(* IEC 61131-3 sources: com.logicals.npe.examples/HIS_Demo/.shadowcopy/src, 6 files *)

(* ---- FB_HISSafety.iecfbd ---- *)
(* Safety FBD template. Two equivalent NC contacts assumed.
   Requires the matching PLCopen Safety library and qualified HIS target setup.
   T#100ms is a DEMO PLACEHOLDER, not a validated discrepancy time.
   Safe communication loss must substitute FALSE at BOTH safe inputs.
   Never replace missing safe input data with standard BOOL simulation values.
   No auto reset or start reset. Reset does not start the process.
*)
FUNCTION_BLOCK FB_HISSafety
  USING safety.plcopen;
VAR_INPUT
    S_EStopA : SAFEBOOL;
    S_EStopB : SAFEBOOL;
    Reset : BOOL;
END_VAR
VAR_OUTPUT
    S_Permit : SAFEBOOL;
    SafetyDemand : BOOL;
    ResetRequest : BOOL;
    Error : BOOL;
    EquivalentDiag : WORD;
    EStopDiag : WORD;
END_VAR
VAR CONSTANT
    S_ResetDisabled : SAFEBOOL := FALSE;
END_VAR
VAR
    fbEquivalent : SF_Equivalent;
    fbEmergencyStop : SF_EmergencyStop;
END_VAR

  (*
    // Network 1: equivalent contacts, emergency stop, diagnostics
    fbEquivalent(Activate := TRUE, S_ChannelA := S_EStopA, S_ChannelB := S_EStopB, DiscrepancyTime := T#100ms);
    fbEmergencyStop(Activate := TRUE, S_EStopIn := fbEquivalent.S_EquivalentOut, S_StartReset := S_ResetDisabled, S_AutoReset := S_ResetDisabled, Reset := Reset, S_EStopOut => S_Permit, SafetyDemand => SafetyDemand, ResetRequest => ResetRequest, DiagCode => EStopDiag);
    EquivalentDiag := fbEquivalent.DiagCode;
    OR(IN1 := fbEquivalent.Error, IN2 := fbEmergencyStop.Error, OR => Error);
  *)

  @C(1) : @FB(fbEquivalent), @R(450.0, 90.0, 360.0, 194.0), @I(@N(Activate), @L(54.5)), @I(@N(S_ChannelA), @L(84.5)), @I(@N(S_ChannelB), @L(114.5)), @I(@N(DiscrepancyTime), @L(144.5)), @O(@N(Ready), @R(54.5)), @O(@N(S_EquivalentOut), @R(84.5)), @O(@N(SafetyDemand), @R(114.5)), @O(@N(Error), @R(144.5)), @O(@N(DiagCode), @R(174.5));
  @C(2) : @FB(fbEmergencyStop), @R(1260.0, 90.0, 360.0, 224.0), @I(@N(Activate), @L(54.5)), @I(@N(S_EStopIn), @L(84.5)), @I(@N(S_StartReset), @L(114.5)), @I(@N(S_AutoReset), @L(144.5)), @I(@N(Reset), @L(174.5)), @O(@N(Ready), @R(54.5)), @O(@N(S_EStopOut), @R(84.5)), @O(@N(SafetyDemand), @R(114.5)), @O(@N(ResetRequest), @R(144.5)), @O(@N(Error), @R(174.5)), @O(@N(DiagCode), @R(204.5));
  @VF(3) : @E(S_EStopA), @R(45.0, 165.0, 300.0, 19.0);
  @VF(4) : @E(S_EStopB), @R(45.0, 195.0, 300.0, 19.0);
  @VF(5) : @E(Reset), @R(870.0, 255.0, 300.0, 19.0);
  @VF(6) : @E(S_Permit), @R(1710.0, 165.0, 300.0, 19.0);
  @VF(7) : @E(SafetyDemand), @R(1710.0, 195.0, 300.0, 19.0);
  @VF(8) : @E(ResetRequest), @R(1710.0, 225.0, 300.0, 19.0);
  @VF(9) : @E(EStopDiag), @R(1710.0, 285.0, 300.0, 19.0);
  @VF(10) : @E(EquivalentDiag), @R(870.0, 375.0, 300.0, 19.0);
  @C(11) : @F(OR), @R(1260.0, 510.0, 180.0, 104.0), BOOL, @I(@N(IN1), @L(54.5)), @I(@N(IN2), @L(84.5)), @O(@N(OR), @R(54.5));
  @VF(12) : @E(Error), @R(1530.0, 555.0, 300.0, 19.0);

  @VF(25) : @E(TRUE), @R(45.0, 135.0, 300.0, 19.0);
  @VF(26) : @E(T#100ms), @R(45.0, 225.0, 300.0, 19.0);
  @VF(27) : @E(TRUE), @R(870.0, 135.0, 300.0, 19.0);
  @VF(28) : @E(S_ResetDisabled), @R(870.0, 195.0, 300.0, 19.0);
  @VF(29) : @E(S_ResetDisabled), @R(870.0, 225.0, 300.0, 19.0);

  @G(13) : @L(@VF(3).o, @C(1).S_ChannelA);
  @G(14) : @L(@VF(4).o, @C(1).S_ChannelB);
  @G(15) : @L(@C(1).S_EquivalentOut, @C(2).S_EStopIn);
  @G(16) : @L(@VF(5).o, @C(2).Reset);
  @G(17) : @L(@C(2).S_EStopOut, @VF(6).i);
  @G(18) : @L(@C(2).SafetyDemand, @VF(7).i);
  @G(19) : @L(@C(2).ResetRequest, @VF(8).i);
  @G(20) : @L(@C(2).DiagCode, @VF(9).i);
  @G(21) : @L(@C(1).DiagCode, @VF(10).i);
  @G(22) : @L(@C(1).Error, @C(11).IN1);
  @G(23) : @L(@C(2).Error, @C(11).IN2);
  @G(24) : @L(@C(11).OR, @VF(12).i);
  @G(30) : @L(@VF(25).o, @C(1).Activate);
  @G(31) : @L(@VF(26).o, @C(1).DiscrepancyTime);
  @G(32) : @L(@VF(27).o, @C(2).Activate);
  @G(33) : @L(@VF(28).o, @C(2).S_StartReset);
  @G(34) : @L(@VF(29).o, @C(2).S_AutoReset);
END_FUNCTION_BLOCK

(* ---- FB_PackagingDataSimulation.iecst ---- *)
(* Simulation-only synthetic process data and harmless demo-load outputs.
 * Called after FB_PackagingLine, only in SimMode. Not a safety function.
 *)
FUNCTION_BLOCK FB_PackagingDataSimulation
    VAR_INPUT
        Reset : BOOL;
        S_Permit : SAFEBOOL;
        S_EStopReleased : SAFEBOOL;
        LineState : UINT;
        LineFault : BOOL;
        CycleDone : BOOL;
        FastCycle : BOOL;
        Heartbeat : BOOL;
    END_VAR
    VAR_OUTPUT
        S_DataPlausible : SAFEBOOL;
    END_VAR
    VAR
        tSecond : TON;
        PrevJam : BOOL;
        PrevGuardClosed : SAFEBOOL := TRUE;
        PrevEStopReleased : SAFEBOOL := FALSE;
        PreviousLineState : UINT;
    END_VAR
    VAR_EXTERNAL
        S_InfeedGuardClosed : SAFEBOOL;
        S_SealingGuardClosed : SAFEBOOL;
        S_OutfeedGuardClosed : SAFEBOOL;
        S_ServiceDoorClosed : SAFEBOOL;
        S_AirSupplyReady : SAFEBOOL;
        S_InfeedZoneStatus : SAFEBYTE;
        S_SealingZoneStatus : SAFEBYTE;
        S_OutfeedZoneStatus : SAFEBYTE;
        S_GuardLockStatus : SAFEBYTE;
        S_SafeDriveStatus : SAFEBYTE;
        S_InfeedDiagnosticCode : SAFEWORD;
        S_SealingDiagnosticCode : SAFEWORD;
        S_OutfeedDiagnosticCode : SAFEWORD;
        S_SafetyBusDiagnosticCode : SAFEWORD;
        S_DriveDiagnosticCode : SAFEWORD;
        S_ZonePermissionMask : SAFEDWORD;
        S_GuardMonitoringMask : SAFEDWORD;
        S_DriveEnableMask : SAFEDWORD;
        S_ActiveSafetyDemandMask : SAFEDWORD;
        S_ConfirmedSafetyDemandMask : SAFEDWORD;
        S_InfeedMotionDirection : SAFESINT;
        S_SealingMotionDirection : SAFESINT;
        S_OutfeedMotionDirection : SAFESINT;
        S_FilmFeedMotionDirection : SAFESINT;
        S_RejectGateMotionDirection : SAFESINT;
        S_SealingTemperatureLimit_dC : SAFEINT;
        S_SealingTemperatureActual_dC : SAFEINT;
        S_AmbientTemperatureActual_dC : SAFEINT;
        S_MinSealingTemperature_dC : SAFEINT;
        S_MaxSealingTemperature_dC : SAFEINT;
        S_InfeedStopPosition_mm : SAFEDINT;
        S_SealingStopPosition_mm : SAFEDINT;
        S_OutfeedStopPosition_mm : SAFEDINT;
        S_CartonTrackingPosition_mm : SAFEDINT;
        S_MaxStoppingDistance_mm : SAFEDINT;
        S_InfeedSensorCount : SAFEUSINT;
        S_SealingSensorCount : SAFEUSINT;
        S_OutfeedSensorCount : SAFEUSINT;
        S_GuardChannelCount : SAFEUSINT;
        S_DriveFeedbackChannelCount : SAFEUSINT;
        S_InfeedSpeedLimit_mm_s : SAFEUINT;
        S_OutfeedSpeedLimit_mm_s : SAFEUINT;
        S_MinAirPressure_mbar : SAFEUINT;
        S_MaxAirPressure_mbar : SAFEUINT;
        S_MotorCurrentLimit_mA : SAFEUINT;
        S_CompletedCartonCount : SAFEUDINT;
        S_RejectedCartonCount : SAFEUDINT;
        S_GuardOpeningCount : SAFEUDINT;
        S_EStopDemandCount : SAFEUDINT;
        S_OperatingTime_s : SAFEUDINT;
        O01 : BOOL;
        O02 : BOOL;
        O03 : BOOL;
        O04 : BOOL;
        O14 : BOOL;
        O15 : BOOL;
        O16 : BOOL;
        O17 : BOOL;
        O18 : BOOL;
        SO01 : SAFEBOOL;
        SO02 : SAFEBOOL;
        SO12 : SAFEBOOL;
        SO13 : SAFEBOOL;
        SO14 : SAFEBOOL;
    END_VAR

    IF Reset THEN
        S_CompletedCartonCount := 0;
        S_RejectedCartonCount := 0;
        S_GuardOpeningCount := 0;
        S_EStopDemandCount := 0;
        S_OperatingTime_s := 0;
        S_SealingTemperatureActual_dC := 1650;
        S_CartonTrackingPosition_mm := 0;
        PrevJam := LineFault;
        PrevGuardClosed := TRUE;
        PrevEStopReleased := S_EStopReleased;
        PreviousLineState := 0;
    END_IF;
    (* Telemetry tick: task-quantised nominal second, not a precision clock. *)
    tSecond(IN := NOT tSecond.Q AND NOT Reset, PT := T#1s);

    S_InfeedGuardClosed := TRUE;
    S_SealingGuardClosed := TRUE;
    S_OutfeedGuardClosed := TRUE;
    S_ServiceDoorClosed := TRUE;
    IF LineFault THEN S_ServiceDoorClosed := FALSE; END_IF;
    S_AirSupplyReady := S_EStopReleased;
    S_SealingTemperatureLimit_dC := 1800;
    S_MinSealingTemperature_dC := 1600;
    S_MaxSealingTemperature_dC := 2000;
    S_AmbientTemperatureActual_dC := 230;
    S_InfeedStopPosition_mm := 1000;
    S_SealingStopPosition_mm := 2000;
    S_OutfeedStopPosition_mm := 3000;
    S_MaxStoppingDistance_mm := 200;
    S_InfeedSpeedLimit_mm_s := 250;
    S_OutfeedSpeedLimit_mm_s := 250;
    IF FastCycle THEN
        S_InfeedSpeedLimit_mm_s := 500;
        S_OutfeedSpeedLimit_mm_s := 500;
    END_IF;
    S_MinAirPressure_mbar := 5500;
    S_MaxAirPressure_mbar := 7500;
    S_MotorCurrentLimit_mA := 4500;
    S_InfeedSensorCount := 2;
    S_SealingSensorCount := 2;
    S_OutfeedSensorCount := 2;
    S_GuardChannelCount := 4;
    S_DriveFeedbackChannelCount := 3;

    (* Zone status 0 blocked, 1 idle, 2 moving, 3 jam. *)
    S_InfeedZoneStatus := 0;
    S_SealingZoneStatus := 0;
    S_OutfeedZoneStatus := 0;
    IF S_Permit AND NOT LineFault THEN
        S_InfeedZoneStatus := 1;
        S_SealingZoneStatus := 1;
        S_OutfeedZoneStatus := 1;
        IF LineState = 20 THEN S_InfeedZoneStatus := 2; END_IF;
        IF LineState = 30 THEN S_SealingZoneStatus := 2; END_IF;
        IF LineState = 40 THEN S_OutfeedZoneStatus := 2; END_IF;
    END_IF;
    IF LineFault THEN S_SealingZoneStatus := 3; END_IF;
    S_GuardLockStatus := 1;
    IF NOT S_ServiceDoorClosed THEN S_GuardLockStatus := 0; END_IF;
    S_SafeDriveStatus := 0;
    IF S_Permit AND S_ServiceDoorClosed THEN S_SafeDriveStatus := 1; END_IF;
    S_InfeedDiagnosticCode := 0;
    S_SealingDiagnosticCode := 0;
    S_OutfeedDiagnosticCode := 0;
    S_SafetyBusDiagnosticCode := 0;
    S_DriveDiagnosticCode := 0;
    IF LineFault THEN S_SealingDiagnosticCode := 16#1001; END_IF;
    IF NOT S_EStopReleased THEN S_SafetyBusDiagnosticCode := 16#2001; END_IF;
    IF NOT S_Permit THEN S_DriveDiagnosticCode := 16#3001; END_IF;

    (* Zones bits 0..2, guards bits 0..3; demand bit 0 E-stop,
       bit 1 virtual service access during jam recovery. *)
    S_ZonePermissionMask := 0;
    IF S_Permit AND S_ServiceDoorClosed AND S_AirSupplyReady THEN S_ZonePermissionMask := 7; END_IF;
    S_GuardMonitoringMask := 15;
    IF NOT S_ServiceDoorClosed THEN S_GuardMonitoringMask := 7; END_IF;
    (* SAFEDWORD is a bitstring, not an arithmetic integer.
       Explicit patterns: bit 0 = E-stop, bit 1 = virtual service door. *)
    S_ActiveSafetyDemandMask := 16#00000000;
    IF NOT S_EStopReleased THEN
        S_ActiveSafetyDemandMask := 16#00000001;
        IF NOT S_ServiceDoorClosed THEN S_ActiveSafetyDemandMask := 16#00000003; END_IF;
    ELSIF NOT S_ServiceDoorClosed THEN
        S_ActiveSafetyDemandMask := 16#00000002;
    END_IF;
    S_ConfirmedSafetyDemandMask := S_ActiveSafetyDemandMask;
    S_DriveEnableMask := 0;
    S_InfeedMotionDirection := 0;
    S_SealingMotionDirection := 0;
    S_OutfeedMotionDirection := 0;
    S_FilmFeedMotionDirection := 0;
    S_RejectGateMotionDirection := 0;
    IF S_ZonePermissionMask = 7 THEN
        IF LineState = 20 THEN S_DriveEnableMask := 1; S_InfeedMotionDirection := 1; END_IF;
        IF LineState = 30 THEN S_DriveEnableMask := 2; S_SealingMotionDirection := 1; S_FilmFeedMotionDirection := 1; END_IF;
        IF LineState = 40 THEN S_DriveEnableMask := 4; S_OutfeedMotionDirection := 1; END_IF;
    END_IF;
    (* Signed virtual sample; no physical motor is commanded in reverse. *)
    IF LineFault THEN S_RejectGateMotionDirection := -1; END_IF;

    IF LineState <> PreviousLineState THEN
        IF LineState = 20 THEN S_CartonTrackingPosition_mm := 0; END_IF;
        IF (LineState = 30) OR (LineState = 40) THEN S_CartonTrackingPosition_mm := S_SealingStopPosition_mm; END_IF;
        IF LineState = 50 THEN S_CartonTrackingPosition_mm := S_OutfeedStopPosition_mm; END_IF;
    END_IF;
    IF (LineState = 0) OR (LineState = 10) THEN S_CartonTrackingPosition_mm := 0; END_IF;
    IF tSecond.Q THEN
        IF S_OperatingTime_s < 1000000000 THEN S_OperatingTime_s := S_OperatingTime_s + 1; END_IF;
        IF S_SealingTemperatureActual_dC < S_SealingTemperatureLimit_dC THEN
            S_SealingTemperatureActual_dC := S_SealingTemperatureActual_dC + 10;
            IF S_SealingTemperatureActual_dC > S_SealingTemperatureLimit_dC THEN S_SealingTemperatureActual_dC := S_SealingTemperatureLimit_dC; END_IF;
        END_IF;
        IF (S_InfeedMotionDirection = 1) AND (S_CartonTrackingPosition_mm < S_InfeedStopPosition_mm) THEN
            S_CartonTrackingPosition_mm := S_CartonTrackingPosition_mm + 250;
            IF S_CartonTrackingPosition_mm > S_InfeedStopPosition_mm THEN S_CartonTrackingPosition_mm := S_InfeedStopPosition_mm; END_IF;
        END_IF;
        IF (S_OutfeedMotionDirection = 1) AND (S_CartonTrackingPosition_mm < S_OutfeedStopPosition_mm) THEN
            S_CartonTrackingPosition_mm := S_CartonTrackingPosition_mm + 250;
            IF S_CartonTrackingPosition_mm > S_OutfeedStopPosition_mm THEN S_CartonTrackingPosition_mm := S_OutfeedStopPosition_mm; END_IF;
        END_IF;
    END_IF;
    (* Separate simulation-session counters, saturated rather than wrapped. *)
    IF NOT Reset THEN
        IF CycleDone AND (S_CompletedCartonCount < 1000000000) THEN S_CompletedCartonCount := S_CompletedCartonCount + 1; END_IF;
        IF LineFault AND NOT PrevJam AND (S_RejectedCartonCount < 1000000000) THEN S_RejectedCartonCount := S_RejectedCartonCount + 1; END_IF;
        IF NOT S_ServiceDoorClosed AND PrevGuardClosed AND (S_GuardOpeningCount < 1000000000) THEN S_GuardOpeningCount := S_GuardOpeningCount + 1; END_IF;
        IF NOT S_EStopReleased AND PrevEStopReleased AND (S_EStopDemandCount < 1000000000) THEN S_EStopDemandCount := S_EStopDemandCount + 1; END_IF;
    END_IF;
    PrevJam := LineFault;
    PrevGuardClosed := S_ServiceDoorClosed;
    PrevEStopReleased := S_EStopReleased;
    PreviousLineState := LineState;

    (* All 50 globals are read in the validity/data chain below. *)
    S_DataPlausible :=
        S_InfeedGuardClosed AND S_SealingGuardClosed AND S_OutfeedGuardClosed
        AND (S_ServiceDoorClosed OR (S_GuardLockStatus = 0))
        AND (S_AirSupplyReady OR (S_ActiveSafetyDemandMask <> 0))
        AND (S_InfeedZoneStatus <= 3) AND (S_SealingZoneStatus <= 3) AND (S_OutfeedZoneStatus <= 3)
        AND (S_GuardLockStatus <= 1) AND (S_SafeDriveStatus <= 1)
        AND (S_InfeedDiagnosticCode = 0) AND ((S_SealingDiagnosticCode = 0) OR (S_SealingDiagnosticCode = 16#1001))
        AND (S_OutfeedDiagnosticCode = 0) AND ((S_SafetyBusDiagnosticCode = 0) OR (S_SafetyBusDiagnosticCode = 16#2001))
        AND ((S_DriveDiagnosticCode = 0) OR (S_DriveDiagnosticCode = 16#3001))
        AND (S_ZonePermissionMask <= 7) AND (S_GuardMonitoringMask <= 15) AND (S_DriveEnableMask <= 7)
        AND (S_ActiveSafetyDemandMask <= 3) AND (S_ConfirmedSafetyDemandMask = S_ActiveSafetyDemandMask)
        AND (S_InfeedMotionDirection >= 0) AND (S_InfeedMotionDirection <= 1)
        AND (S_SealingMotionDirection >= 0) AND (S_SealingMotionDirection <= 1)
        AND (S_OutfeedMotionDirection >= 0) AND (S_OutfeedMotionDirection <= 1)
        AND (S_FilmFeedMotionDirection >= 0) AND (S_FilmFeedMotionDirection <= 1)
        AND (S_RejectGateMotionDirection >= -1) AND (S_RejectGateMotionDirection <= 0)
        AND (S_SealingTemperatureLimit_dC >= S_MinSealingTemperature_dC)
        AND (S_SealingTemperatureLimit_dC <= S_MaxSealingTemperature_dC)
        AND (S_SealingTemperatureActual_dC >= S_MinSealingTemperature_dC)
        AND (S_SealingTemperatureActual_dC <= S_MaxSealingTemperature_dC)
        AND (S_AmbientTemperatureActual_dC >= 0) AND (S_AmbientTemperatureActual_dC <= 500)
        AND (S_InfeedStopPosition_mm > S_MaxStoppingDistance_mm)
        AND (S_SealingStopPosition_mm > S_InfeedStopPosition_mm)
        AND (S_OutfeedStopPosition_mm > S_SealingStopPosition_mm)
        AND (S_CartonTrackingPosition_mm >= 0) AND (S_CartonTrackingPosition_mm <= S_OutfeedStopPosition_mm)
        AND (S_InfeedSensorCount = 2) AND (S_SealingSensorCount = 2) AND (S_OutfeedSensorCount = 2)
        AND (S_GuardChannelCount = 4) AND (S_DriveFeedbackChannelCount = 3)
        AND (S_InfeedSpeedLimit_mm_s > 0) AND (S_InfeedSpeedLimit_mm_s <= 500)
        AND (S_OutfeedSpeedLimit_mm_s > 0) AND (S_OutfeedSpeedLimit_mm_s <= 500)
        AND (S_MinAirPressure_mbar < S_MaxAirPressure_mbar) AND (S_MotorCurrentLimit_mA > 0)
        AND (S_CompletedCartonCount <= 1000000000) AND (S_RejectedCartonCount <= 1000000000)
        AND (S_GuardOpeningCount = S_RejectedCartonCount)
        AND (S_EStopDemandCount <= 1000000000) AND (S_OperatingTime_s <= 1000000000);

    O01 := S_Permit AND S_DataPlausible AND (S_InfeedMotionDirection = 1);
    O02 := S_Permit AND S_DataPlausible AND (S_SealingMotionDirection = 1);
    O03 := S_Permit AND S_DataPlausible AND (S_OutfeedMotionDirection = 1);
    O04 := S_Permit AND S_DataPlausible AND (S_FilmFeedMotionDirection = 1);
    O14 := S_Permit AND S_DataPlausible AND (S_ZonePermissionMask = 7);
    O15 := S_Permit AND S_DataPlausible AND Heartbeat;
    O16 := S_Permit AND S_DataPlausible AND (S_SealingDiagnosticCode <> 0);
    O17 := S_Permit AND S_DataPlausible AND (S_SealingTemperatureActual_dC >= S_SealingTemperatureLimit_dC);
    O18 := S_Permit AND S_DataPlausible AND (S_GuardMonitoringMask = 15);
    (* Safe-typed expressions; demo indications, not validated safety outputs. *)
    SO01 := S_Permit AND S_DataPlausible AND S_AirSupplyReady;
    SO02 := S_Permit AND S_DataPlausible AND S_ServiceDoorClosed;
    SO12 := S_Permit AND S_DataPlausible AND S_InfeedGuardClosed AND (S_InfeedMotionDirection = 1);
    SO13 := S_Permit AND S_DataPlausible AND S_SealingGuardClosed AND (S_SealingMotionDirection = 1);
    SO14 := S_Permit AND S_DataPlausible AND S_OutfeedGuardClosed AND (S_OutfeedMotionDirection = 1);
END_FUNCTION_BLOCK

(* ---- FB_PackagingIndicators.iecfbd ---- *)
(* Non-safety FBD. Suggested four standard LED functions.
   All physical output assignments remain open.
*)
FUNCTION_BLOCK FB_PackagingIndicators
VAR_INPUT
    Permit : BOOL;
    Ready : BOOL;
    Infeed : BOOL;
    Sealing : BOOL;
    Outfeed : BOOL;
    Complete : BOOL;
    Blocked : BOOL;
    ProcessFault : BOOL;
    SafetyError : BOOL;
    ResetRequest : BOOL;
    Heartbeat : BOOL;
END_VAR
VAR_OUTPUT
    LedReady : BOOL;
    LedConveyor : BOOL;
    LedSealing : BOOL;
    LedAttention : BOOL;
END_VAR

  (*
    Explicit Boolean gates; value fields contain single variables only.
    OR(IN1 := Ready, IN2 := Complete);
    AND(IN1 := Permit, IN2 := @C(1).OR);
    OR(IN1 := Infeed, IN2 := Outfeed);
    AND(IN1 := Permit, IN2 := @C(7).OR, IN3 := Heartbeat);
    AND(IN1 := Permit, IN2 := Sealing, IN3 := Heartbeat);
    NOT(IN := ResetRequest);
    AND(IN1 := Blocked, IN2 := @C(19).NOT);
    AND(IN1 := ResetRequest, IN2 := Heartbeat);
    OR(IN1 := @C(21).AND, IN2 := ProcessFault, IN3 := SafetyError, IN4 := @C(23).AND);
  *)

  @C(1) : @F(OR), @R(390.0, 90.0, 180.0, 104.0), BOOL, @I(@N(IN1), @L(54.5)), @I(@N(IN2), @L(84.5)), @O(@N(OR), @R(54.5));
  @VF(2) : @E(Ready), @R(45.0, 135.0, 180.0, 19.0);
  @VF(3) : @E(Complete), @R(45.0, 165.0, 180.0, 19.0);
  @C(4) : @F(AND), @R(900.0, 60.0, 180.0, 104.0), BOOL, @I(@N(IN1), @L(54.5)), @I(@N(IN2), @L(84.5)), @O(@N(AND), @R(54.5));
  @VF(5) : @E(Permit), @R(645.0, 105.0, 180.0, 19.0);
  @VF(6) : @E(LedReady), @R(1230.0, 105.0, 180.0, 19.0);
  @C(7) : @F(OR), @R(390.0, 390.0, 180.0, 104.0), BOOL, @I(@N(IN1), @L(54.5)), @I(@N(IN2), @L(84.5)), @O(@N(OR), @R(54.5));
  @VF(8) : @E(Infeed), @R(45.0, 435.0, 180.0, 19.0);
  @VF(9) : @E(Outfeed), @R(45.0, 465.0, 180.0, 19.0);
  @C(10) : @F(AND), @R(900.0, 360.0, 180.0, 134.0), BOOL, @I(@N(IN1), @L(54.5)), @I(@N(IN2), @L(84.5)), @I(@N(IN3), @L(114.5)), @O(@N(AND), @R(54.5));
  @VF(11) : @E(Permit), @R(645.0, 405.0, 180.0, 19.0);
  @VF(12) : @E(Heartbeat), @R(645.0, 465.0, 180.0, 19.0);
  @VF(13) : @E(LedConveyor), @R(1230.0, 405.0, 180.0, 19.0);
  @C(14) : @F(AND), @R(900.0, 660.0, 180.0, 134.0), BOOL, @I(@N(IN1), @L(54.5)), @I(@N(IN2), @L(84.5)), @I(@N(IN3), @L(114.5)), @O(@N(AND), @R(54.5));
  @VF(15) : @E(Permit), @R(645.0, 705.0, 180.0, 19.0);
  @VF(16) : @E(Sealing), @R(645.0, 735.0, 180.0, 19.0);
  @VF(17) : @E(Heartbeat), @R(645.0, 765.0, 180.0, 19.0);
  @VF(18) : @E(LedSealing), @R(1230.0, 705.0, 180.0, 19.0);
  @C(19) : @F(NOT), @R(375.0, 1080.0, 180.0, 74.0), BOOL, @I(@N(IN), @L(54.5)), @O(@N(NOT), @R(54.5));
  @VF(20) : @E(ResetRequest), @R(45.0, 1125.0, 180.0, 19.0);
  @C(21) : @F(AND), @R(660.0, 1050.0, 180.0, 104.0), BOOL, @I(@N(IN1), @L(54.5)), @I(@N(IN2), @L(84.5)), @O(@N(AND), @R(54.5));
  @VF(22) : @E(Blocked), @R(375.0, 1035.0, 180.0, 19.0);
  @C(23) : @F(AND), @R(660.0, 1230.0, 180.0, 104.0), BOOL, @I(@N(IN1), @L(54.5)), @I(@N(IN2), @L(84.5)), @O(@N(AND), @R(54.5));
  @VF(24) : @E(ResetRequest), @R(375.0, 1275.0, 180.0, 19.0);
  @VF(25) : @E(Heartbeat), @R(375.0, 1305.0, 180.0, 19.0);
  @C(26) : @F(OR), @R(1200.0, 1050.0, 180.0, 164.0), BOOL, @I(@N(IN1), @L(54.5)), @I(@N(IN2), @L(84.5)), @I(@N(IN3), @L(114.5)), @I(@N(IN4), @L(144.5)), @O(@N(OR), @R(54.5));
  @VF(27) : @E(ProcessFault), @R(930.0, 1125.0, 180.0, 19.0);
  @VF(28) : @E(SafetyError), @R(930.0, 1155.0, 180.0, 19.0);
  @VF(29) : @E(LedAttention), @R(1500.0, 1095.0, 180.0, 19.0);

  @G(30) : @L(@VF(2).o, @C(1).IN1);
  @G(31) : @L(@VF(3).o, @C(1).IN2);
  @G(32) : @L(@VF(5).o, @C(4).IN1);
  @G(33) : @L(@C(1).OR, @C(4).IN2);
  @G(34) : @L(@C(4).AND, @VF(6).i);
  @G(35) : @L(@VF(8).o, @C(7).IN1);
  @G(36) : @L(@VF(9).o, @C(7).IN2);
  @G(37) : @L(@VF(11).o, @C(10).IN1);
  @G(38) : @L(@C(7).OR, @C(10).IN2);
  @G(39) : @L(@VF(12).o, @C(10).IN3);
  @G(40) : @L(@C(10).AND, @VF(13).i);
  @G(41) : @L(@VF(15).o, @C(14).IN1);
  @G(42) : @L(@VF(16).o, @C(14).IN2);
  @G(43) : @L(@VF(17).o, @C(14).IN3);
  @G(44) : @L(@C(14).AND, @VF(18).i);
  @G(45) : @L(@VF(20).o, @C(19).IN);
  @G(46) : @L(@VF(22).o, @C(21).IN1);
  @G(47) : @L(@C(19).NOT, @C(21).IN2);
  @G(48) : @L(@VF(24).o, @C(23).IN1);
  @G(49) : @L(@VF(25).o, @C(23).IN2);
  @G(50) : @L(@C(21).AND, @C(26).IN1);
  @G(51) : @L(@VF(27).o, @C(26).IN2);
  @G(52) : @L(@VF(28).o, @C(26).IN3);
  @G(53) : @L(@C(23).AND, @C(26).IN4);
  @G(54) : @L(@C(26).OR, @VF(29).i);
END_FUNCTION_BLOCK

(* ---- FB_PackagingLine.iecst ---- *)
(* HIS Packaging Line / SPS 2026
 *    Non-safety simulation. Never use these outputs as a safety function.
 *    Call once per cyclic task. No physical I/O addresses are assigned.
 *)
FUNCTION_BLOCK FB_PackagingLine
	VAR_INPUT
		Enable : BOOL;
		Permit : BOOL; (* Read-only status copy from the safety POU. *)
		Start : BOOL;
		Stop : BOOL;
		FastCycle : BOOL;
		Jam : BOOL; (* Simulated carton jam, NOT a safety fault. *)
		AckJam : BOOL;
	END_VAR
	VAR_OUTPUT
		State : UINT;
		(* 0 blocked, 10 ready, 20 infeed, 30 sealing,
		 40 outfeed, 50 complete, 90 carton jam *)
		Ready : BOOL;
		Infeed : BOOL;
		Sealing : BOOL;
		Outfeed : BOOL;
		Complete : BOOL;
		Blocked : BOOL;
		Fault : BOOL;
		Running : BOOL;
		Heartbeat : BOOL;
		CycleDone : BOOL; (* One scan pulse after carton leaves station. *)
		CartonsPacked : UDINT;
		FastCycleActive : BOOL;
	END_VAR
	VAR
		PrevStart : BOOL;
		PrevAck : BOOL;
		FirstScan : BOOL := TRUE;
		StartEdge : BOOL;
		AckEdge : BOOL;
		StartArmed : BOOL;
		FaultLatched : BOOL;
		InfeedTime : TIME := T#3s;
		SealTime : TIME := T#2s;
		OutfeedTime : TIME := T#2s;
		tInfeed : TON;
		tSeal : TON;
		tOutfeed : TON;
		tSuccess : TON;
		tBlink : TON;
	END_VAR

	(* Suppress edges on startup; held Start never causes a restart. *)
	StartEdge := Start AND NOT PrevStart AND NOT FirstScan;
	AckEdge := AckJam AND NOT PrevAck AND NOT FirstScan;
	PrevStart := Start;
	PrevAck := AckJam;
	FirstScan := FALSE;
	CycleDone := FALSE;

	(* Timers are executed on every scan, also when disabled. *)
	tBlink(IN := NOT tBlink.Q, PT := T#250ms);
	IF tBlink.Q THEN
		Heartbeat := NOT Heartbeat;
	END_IF;
	tInfeed(IN := (State = 20) AND Enable AND Permit AND NOT Stop
            AND NOT Jam, PT := InfeedTime);
	tSeal(IN := (State = 30) AND Enable AND Permit AND NOT Stop
             AND NOT Jam, PT := SealTime);
	tOutfeed(IN := (State = 40) AND Enable AND Permit AND NOT Stop
              AND NOT Jam, PT := OutfeedTime);
	tSuccess(IN := (State = 50) AND Enable AND Permit AND NOT Stop
               AND NOT Jam, PT := T#1s);

	(* Keep process faults latched even across a safety interruption. *)
	IF Jam AND Enable AND Permit
   AND ((State = 20) OR (State = 30) OR (State = 40)) THEN
		FaultLatched := TRUE;
	END_IF;
	IF AckEdge AND NOT Jam AND Enable AND Permit THEN
		FaultLatched := FALSE;
	END_IF;

	(* Priority: no permit / disabled > process fault > stop > sequence. *)
	IF NOT Enable OR NOT Permit THEN
		State := 0;

		FastCycleActive := FALSE;
		StartArmed := FALSE;
	ELSIF FaultLatched THEN
		State := 90;

		FastCycleActive := FALSE;
		StartArmed := FALSE;
	ELSIF Stop THEN
		State := 10;

		FastCycleActive := FALSE;
		StartArmed := FALSE;
	ELSE
		CASE State OF
			0, 90:
			State := 10;

			FastCycleActive := FALSE;
			StartArmed := FALSE;
			10:
            IF NOT Start THEN
				StartArmed := TRUE;
			END_IF;
			IF StartEdge AND StartArmed AND NOT Jam
               AND NOT AckJam THEN
				FastCycleActive := FastCycle; (* Latch throughput mode for this carton. *)
				IF FastCycleActive THEN
					InfeedTime := T#1500ms;
					SealTime := T#1s;
					OutfeedTime := T#1s;
				ELSE
					InfeedTime := T#3s;
					SealTime := T#2s;
					OutfeedTime := T#2s;
				END_IF;
				StartArmed := FALSE;

				State := 20;
			END_IF;
			20:
            IF tInfeed.Q THEN
				State := 30;
			END_IF;
			30:
            IF tSeal.Q THEN

				State := 40;
			END_IF;
			40:
            IF tOutfeed.Q THEN
				IF CartonsPacked < UDINT#4294967295 THEN
					CartonsPacked := CartonsPacked + 1;
				END_IF;
				CycleDone := TRUE;
				State := 50;
			END_IF;
			50:
            IF tSuccess.Q THEN
				State := 10;
				FastCycleActive := FALSE;
				StartArmed := FALSE;
			END_IF;
		ELSE
			FaultLatched := TRUE;
			State := 90;

			FastCycleActive := FALSE;
			StartArmed := FALSE;
		END_CASE;
	END_IF;

	Blocked := NOT Enable OR NOT Permit;
	Fault := FaultLatched;
	Ready := (State = 10) AND Enable AND Permit AND NOT FaultLatched
         AND NOT Stop AND NOT Jam AND NOT AckJam;
	Infeed := State = 20;
	Sealing := State = 30;
	Outfeed := State = 40;
	Complete := State = 50;
	Running := Infeed OR Sealing OR Outfeed;
END_FUNCTION_BLOCK

(* ---- FB_PackagingSimulation.iecst ---- *)
(* Automatic exhibition simulation; not a physical safety input source.
 * Called ONLY while PRG_HISDemo.SimMode is TRUE.
 * Drives simulated commands through the unchanged safety/process blocks.
 * Reset on every mode entry; feedback comes from the previous program scan.
 *)
FUNCTION_BLOCK FB_PackagingSimulation
    VAR_INPUT
        Reset : BOOL;
        Permit : BOOL;
        LineReady : BOOL;
        LineState : UINT;
        LineFault : BOOL;
        InjectFaults : BOOL;
        FastCycle : BOOL;
    END_VAR
    VAR_OUTPUT
        EStopReleased : SAFEBOOL;
        Enable : BOOL;
        Start : BOOL;
        Stop : BOOL;
        SafetyReset : BOOL;
        Jam : BOOL;
        AckJam : BOOL;
        FastCycleCommand : BOOL;
        (* 0 boot; 10 release; 20 reset gap; 30 reset pulse; 40 ready;
           50 start pulse; 60 packaging; 70 jam; 80 clear jam;
           90 acknowledge; 100 emergency stop. *)
        State : UINT;
        AttemptInRound : UINT;
        (* 0 none; 1 normal carton; 2 jam demonstration; 3 E-stop demonstration. *)
        Scenario : UINT;
    END_VAR
    VAR
        tBoot : TON;
        tRelease : TON;
        tResetGap : TON;
        tResetPulse : TON;
        tReady : TON;
        tStart : TON;
        tJam : TON;
        tJamClear : TON;
        tAck : TON;
        tEStop : TON;
    END_VAR

    IF Reset THEN
        State := 0;
        AttemptInRound := 0;
        Scenario := 0;
    END_IF;

    (* Separate timers ensure every phase receives a fresh interval.
       Reset also clears timers left active when the block was not called. *)
    tBoot(IN := (State = 0) AND NOT Reset, PT := T#1s);
    tRelease(IN := (State = 10) AND NOT Reset, PT := T#1s);
    tResetGap(IN := (State = 20) AND NOT Reset, PT := T#500ms);
    tResetPulse(IN := (State = 30) AND NOT Reset, PT := T#500ms);
    tReady(IN := (State = 40) AND LineReady AND Permit AND NOT Reset, PT := T#500ms);
    tStart(IN := (State = 50) AND NOT Reset, PT := T#500ms);
    tJam(IN := (State = 70) AND NOT Reset, PT := T#3s);
    tJamClear(IN := (State = 80) AND NOT Reset, PT := T#500ms);
    tAck(IN := (State = 90) AND NOT Reset, PT := T#500ms);
    tEStop(IN := (State = 100) AND NOT Reset, PT := T#3s);

    IF NOT Reset THEN
        CASE State OF
            0:
                IF tBoot.Q THEN State := 10; END_IF;
            10:
                IF tRelease.Q THEN State := 20; END_IF;
            20:
                IF Permit THEN
                    IF LineFault THEN State := 80; ELSE State := 40; END_IF;
                ELSIF tResetGap.Q THEN
                    State := 30;
                END_IF;
            30:
                IF tResetPulse.Q THEN
                    IF Permit THEN
                        IF LineFault THEN State := 80; ELSE State := 40; END_IF;
                    ELSE
                        State := 20;
                    END_IF;
                END_IF;
            40:
                IF NOT Permit THEN
                    State := 10;
                ELSIF LineFault THEN
                    State := 80;
                ELSIF tReady.Q THEN
                    IF AttemptInRound >= 6 THEN AttemptInRound := 0; END_IF;
                    AttemptInRound := AttemptInRound + 1;
                    Scenario := 1;
                    IF InjectFaults AND (AttemptInRound = 3) THEN Scenario := 2; END_IF;
                    IF InjectFaults AND (AttemptInRound = 6) THEN Scenario := 3; END_IF;
                    State := 50;
                END_IF;
            50:
                IF NOT Permit THEN
                    State := 10;
                ELSIF tStart.Q THEN
                    State := 60;
                END_IF;
            60:
                IF NOT Permit THEN
                    State := 10;
                ELSIF LineFault THEN
                    State := 80;
                ELSIF (Scenario = 2) AND (LineState = 30) THEN
                    State := 70;
                ELSIF (Scenario = 3) AND (LineState = 30) THEN
                    State := 100;
                ELSIF (LineState = 50) OR LineReady THEN
                    State := 40;
                END_IF;
            70:
                IF tJam.Q THEN State := 80; END_IF;
            80:
                IF NOT Permit THEN
                    State := 10;
                ELSIF tJamClear.Q THEN
                    State := 90;
                END_IF;
            90:
                IF NOT Permit THEN
                    State := 10;
                ELSIF tAck.Q THEN
                    IF LineFault THEN State := 80; ELSE State := 40; END_IF;
                END_IF;
            100:
                IF tEStop.Q THEN State := 10; END_IF;
        ELSE
            State := 0;
            Scenario := 0;
        END_CASE;
    END_IF;

    (* Defined outputs every scan. Both virtual contacts are mapped together
       by the calling program; the PLCopen permit is never forced here. *)
    EStopReleased := FALSE;
    IF (State <> 0) AND (State <> 100) THEN EStopReleased := TRUE; END_IF;
    Enable := State <> 0;
    Start := State = 50;
    Stop := FALSE;
    SafetyReset := State = 30;
    Jam := State = 70;
    AckJam := State = 90;
    FastCycleCommand := FastCycle;
END_FUNCTION_BLOCK

(* ---- PRG_HISDemo.iecst ---- *)
(* HIS Packaging Demo: hardware operation or automatic exhibition simulation.
 * SimMode defaults to FALSE. Simulation ignores the four physical inputs.
 * Only the demo inputs/commands are substituted; PLCopen blocks stay active.
 * Intended for this indicator-only demonstrator, not real actuator operation.
 *)
PROGRAM PRG_HISDemo
	VAR
		SimMode : BOOL := FALSE; (* TRUE = autonomous simulation; FALSE = physical inputs. *)
		SimInjectFaults : BOOL := TRUE; (* Jam on attempt 3, E-stop on attempt 6. *)
		SimFastCycle : BOOL := FALSE;
		SimModePrev : BOOL := FALSE;
		ModeChanged : BOOL;
		HardwareCommandsArmed : BOOL := TRUE;
		Simulation : FB_PackagingSimulation;
		DataSimulation : FB_PackagingDataSimulation;
		SimDataOutputsOwned : BOOL := FALSE;
		(* Selected E-stop input: FALSE = pressed; TRUE = released.
		 Derived every scan from hardware or the simulation block. *)
		Sim_EStopReleased : SAFEBOOL := FALSE;
		(* Derived virtual contacts, overwritten every scan; do not edit online. *)
		S_EStopA : SAFEBOOL;
		S_EStopB : SAFEBOOL;

		CmdEnable : BOOL; (* Latched enable: physical button toggles on each rising edge. *)
		EnableButtonPrev : BOOL := FALSE;
		EnableButtonFirstScan : BOOL := TRUE;
		CmdStart : BOOL;
		CmdStop : BOOL;
		CmdFastCycle : BOOL;
		CmdJam : BOOL;
		CmdSafetyReset : BOOL;
		CmdAckJam : BOOL;

		(* Symbolic outputs: actual terminals will be assigned later. *)
		S_DemoEnable : SAFEBOOL; (* Safe permission indicator; not a run command. *)
		LedReady : BOOL;
		LedConveyor : BOOL;
		LedSealing : BOOL;
		LedAttention : BOOL;

		Safety : FB_HISSafety;
		Line : FB_PackagingLine;
		Lamps : FB_PackagingIndicators;
	END_VAR

	VAR_EXTERNAL
		EStop : SAFEBOOL;
		Button1Input : BOOL;
		Button2Input : BOOL;
		Button3Input : BOOL;
		Button1Indicator : BOOL { description := "��e";
		comment := "Indicator light of first button";};
		Button2Indicator : BOOL { description := "��e";
		comment := "Indicator light of second button";};
		Button3Indicator : BOOL { description := "��e";
		comment := "Indicator light of third button";};
		O01 : BOOL;
		O02 : BOOL;
		O03 : BOOL;
		O04 : BOOL;
		O14 : BOOL;
		O15 : BOOL;
		O16 : BOOL;
		O17 : BOOL;
		O18 : BOOL;
		SO01 : SAFEBOOL;
		SO02 : SAFEBOOL;
		SO12 : SAFEBOOL;
		SO13 : SAFEBOOL;
		SO14 : SAFEBOOL;
	END_VAR

	(* Returning to hardware always requires a new enable/start action.
	   Ignore a held physical enable button during the transition. *)
	ModeChanged := SimMode <> SimModePrev;
	IF ModeChanged THEN
		CmdEnable := FALSE;
		CmdStart := FALSE;
		CmdSafetyReset := FALSE;
		CmdStop := FALSE;
		CmdFastCycle := FALSE;
		CmdJam := FALSE;
		CmdAckJam := FALSE;
		EnableButtonFirstScan := TRUE;
		HardwareCommandsArmed := FALSE;
	END_IF;

	IF SimMode THEN
		(* No physical input is read in this branch. Feedback is one scan old. *)
		Simulation(Reset := ModeChanged, Permit := Safety.S_Permit,
			LineReady := Line.Ready, LineState := Line.State, LineFault := Line.Fault,
			InjectFaults := SimInjectFaults, FastCycle := SimFastCycle);
		Sim_EStopReleased := Simulation.EStopReleased;
		CmdEnable := Simulation.Enable;
		CmdStart := Simulation.Start;
		CmdSafetyReset := Simulation.SafetyReset;
		CmdStop := Simulation.Stop;
		CmdFastCycle := Simulation.FastCycleCommand;
		CmdJam := Simulation.Jam;
		CmdAckJam := Simulation.AckJam;
	ELSE
		Sim_EStopReleased := EStop;
		(* One scan with no E-stop permit on mode exit resets the safety path.
		   Hardware reset/start buttons must also be released before reuse. *)
		IF ModeChanged THEN Sim_EStopReleased := FALSE; END_IF;
		IF Button1Input AND NOT EnableButtonPrev AND NOT EnableButtonFirstScan THEN
			CmdEnable := NOT CmdEnable;
		END_IF;
		EnableButtonPrev := Button1Input;
		EnableButtonFirstScan := FALSE;
		IF NOT ModeChanged AND NOT Button2Input AND NOT Button3Input THEN
			HardwareCommandsArmed := TRUE;
		END_IF;
		CmdSafetyReset := Button2Input AND HardwareCommandsArmed AND NOT ModeChanged;
		CmdStart := Button3Input AND HardwareCommandsArmed AND NOT ModeChanged;
	END_IF;
	SimModePrev := SimMode;

	(* Update both virtual contacts before evaluating safety. *)
	S_EStopA :=	Sim_EStopReleased;
	S_EStopB := Sim_EStopReleased;

	(* Order matters: simulated inputs -> safety -> process -> indication. *)
	Safety(S_EStopA := S_EStopA, S_EStopB := S_EStopB, Reset := CmdSafetyReset);

	(* Safety path does not depend on the standard sequence or standard lamps. *)
	S_DemoEnable := Safety.S_Permit;

	Line(Enable := CmdEnable, Permit := Safety.S_Permit, Start := CmdStart, Stop := CmdStop, FastCycle := CmdFastCycle, Jam := CmdJam, AckJam := CmdAckJam);

    IF SimMode THEN
        DataSimulation(Reset := ModeChanged, S_Permit := Safety.S_Permit,
            S_EStopReleased := Sim_EStopReleased, LineState := Line.State,
            LineFault := Line.Fault, CycleDone := Line.CycleDone,
            FastCycle := Line.FastCycleActive, Heartbeat := Line.Heartbeat);
        SimDataOutputsOwned := TRUE;
    ELSIF SimDataOutputsOwned THEN
        (* One-time mode-exit cleanup. No cyclic hardware-mode writer. *)
        O01 := FALSE;
        O02 := FALSE;
        O03 := FALSE;
        O04 := FALSE;
        O14 := FALSE;
        O15 := FALSE;
        O16 := FALSE;
        O17 := FALSE;
        O18 := FALSE;
        SO01 := FALSE;
        SO02 := FALSE;
        SO12 := FALSE;
        SO13 := FALSE;
        SO14 := FALSE;
        SimDataOutputsOwned := FALSE;
    END_IF;

	Lamps(Permit := Safety.S_Permit, Ready := Line.Ready, Infeed := Line.Infeed, Sealing := Line.Sealing, Outfeed := Line.Outfeed, Complete := Line.Complete, Blocked := Line.Blocked, ProcessFault := Line.Fault, SafetyError := Safety.Error, ResetRequest := Safety.ResetRequest, Heartbeat := Line.Heartbeat, LedReady => LedReady, LedConveyor => LedConveyor, LedSealing => LedSealing, LedAttention => LedAttention);

	Button1Indicator := Lamps.LedReady;
	Button2Indicator := Lamps.LedConveyor;
	Button3Indicator := Lamps.LedSealing;

END_PROGRAM
